(* IEC 61131-3 sources: plc-st-coding-agent/progress/evidence/f14_v2_public_20261112b/jobs/codex_deepseek-v4pro, 5 files *)

(* ---- public-easy-01.candidate_01.st ---- *)
FUNCTION_BLOCK FillingLineControl
VAR_INPUT
    bottleSensor : BOOL;
    cleaningConfirmButton : BOOL;
    fillingConfirmButton : BOOL;
    cappingConfirmButton : BOOL;
    packingConfirmButton : BOOL;
    finishedButton : BOOL;
END_VAR
VAR_OUTPUT
    Pump_Motor : BOOL;
    Filling_Valve : BOOL;
    Capping_Machine : BOOL;
    Packing_Machine : BOOL;
    Completion_Light : BOOL;
END_VAR
VAR
    step : INT := 0;
END_VAR

CASE step OF
    0:
        IF bottleSensor THEN
            step := 1;
        END_IF;

    1:
        IF cleaningConfirmButton THEN
            step := 2;
        END_IF;

    2:
        IF fillingConfirmButton THEN
            step := 3;
        END_IF;

    3:
        IF cappingConfirmButton THEN
            step := 4;
        END_IF;

    4:
        IF packingConfirmButton THEN
            step := 5;
        END_IF;

    5:
        IF finishedButton THEN
            step := 0;
        END_IF;
END_CASE;

Pump_Motor := (step = 1);
Filling_Valve := (step = 2);
Capping_Machine := (step = 3);
Packing_Machine := (step = 4);
Completion_Light := (step = 5);

END_FUNCTION_BLOCK

(* ---- public-easy-02.candidate_01.st ---- *)
FUNCTION_BLOCK FB
VAR_INPUT
    value : DWORD;
END_VAR
VAR_OUTPUT
    hasChanged : BOOL;
    hasRisingEdges : BOOL;
    risingBits : DWORD;
    noOfRisingBits : USINT;
    hasFallingEdges : BOOL;
    fallingBits : DWORD;
    noOfFallingBits : USINT;
END_VAR
VAR
    lastValue : DWORD;
    firstCycle : BOOL := TRUE;
    bitMask : DWORD;
    bitIndex : INT;
END_VAR

noOfRisingBits := USINT#0;
noOfFallingBits := USINT#0;

IF firstCycle THEN
    lastValue := value;
    firstCycle := FALSE;
    hasChanged := FALSE;
    hasRisingEdges := FALSE;
    risingBits := DWORD#0;
    hasFallingEdges := FALSE;
    fallingBits := DWORD#0;
ELSE
    hasChanged := (lastValue <> value);
    risingBits := (NOT lastValue) AND value;
    fallingBits := lastValue AND (NOT value);

    hasRisingEdges := (risingBits <> DWORD#0);
    hasFallingEdges := (fallingBits <> DWORD#0);

    FOR bitIndex := 0 TO 31 DO
        bitMask := SHL(DWORD#1, bitIndex);
        IF ((risingBits AND bitMask) <> DWORD#0) THEN
            noOfRisingBits := noOfRisingBits + USINT#1;
        END_IF;
        IF ((fallingBits AND bitMask) <> DWORD#0) THEN
            noOfFallingBits := noOfFallingBits + USINT#1;
        END_IF;
    END_FOR;

    lastValue := value;
END_IF;

END_FUNCTION_BLOCK

(* ---- public-easy-02.candidate_02.st ---- *)
FUNCTION_BLOCK FB
VAR_INPUT
    value : DWORD;
END_VAR
VAR_OUTPUT
    hasChanged : BOOL;
    hasRisingEdges : BOOL;
    risingBits : DWORD;
    noOfRisingBits : USINT;
    hasFallingEdges : BOOL;
    fallingBits : DWORD;
    noOfFallingBits : USINT;
END_VAR
VAR
    lastValue : DWORD;
    bitIndex : INT;
END_VAR

risingBits := (NOT lastValue) AND value;
fallingBits := lastValue AND (NOT value);

hasChanged := lastValue <> value;
hasRisingEdges := risingBits <> DWORD#0;
hasFallingEdges := fallingBits <> DWORD#0;

noOfRisingBits := USINT#0;
noOfFallingBits := USINT#0;

FOR bitIndex := 0 TO 31 DO
    IF ((SHR(risingBits, bitIndex) AND DWORD#1) <> DWORD#0) THEN
        noOfRisingBits := noOfRisingBits + USINT#1;
    END_IF;

    IF ((SHR(fallingBits, bitIndex) AND DWORD#1) <> DWORD#0) THEN
        noOfFallingBits := noOfFallingBits + USINT#1;
    END_IF;
END_FOR;

lastValue := value;

END_FUNCTION_BLOCK

(* ---- public-easy-03.candidate_01.st ---- *)
FUNCTION_BLOCK AlarmHandling
VAR_INPUT
    Value : REAL;
    hiLevel : REAL;
    loLevel : REAL;
    hystWindow : REAL;
END_VAR

VAR_OUTPUT
    hiAlarm : BOOL;
    loAlarm : BOOL;
    error : BOOL;
    status : WORD;
END_VAR

VAR
    hiAlarmState : BOOL;
    loAlarmState : BOOL;
END_VAR

BEGIN
    hiAlarm := FALSE;
    loAlarm := FALSE;
    error := FALSE;
    status := 16#0000;

    IF loLevel >= hiLevel THEN
        error := TRUE;
        status := 16#8001;
        RETURN;
    END_IF;

    IF hystWindow >= (hiLevel - loLevel) THEN
        error := TRUE;
        status := 16#8002;
        RETURN;
    END_IF;

    IF Value > hiLevel THEN
        hiAlarmState := TRUE;
    ELSIF Value < (hiLevel - hystWindow) THEN
        hiAlarmState := FALSE;
    END_IF;

    IF Value < loLevel THEN
        loAlarmState := TRUE;
    ELSIF Value > (loLevel + hystWindow) THEN
        loAlarmState := FALSE;
    END_IF;

    hiAlarm := hiAlarmState;
    loAlarm := loAlarmState;
END_FUNCTION_BLOCK

(* ---- public-easy-03.candidate_02.st ---- *)
FUNCTION_BLOCK AlarmHandling
VAR_INPUT
    Value : REAL;
    hiLevel : REAL;
    loLevel : REAL;
    hystWindow : REAL;
END_VAR

VAR_OUTPUT
    hiAlarm : BOOL;
    loAlarm : BOOL;
    error : BOOL;
    status : WORD;
END_VAR

BEGIN
    error := FALSE;
    status := WORD#16#0000;

    IF loLevel >= hiLevel THEN
        hiAlarm := FALSE;
        loAlarm := FALSE;
        error := TRUE;
        status := WORD#16#8001;
    ELSIF hystWindow >= (hiLevel - loLevel) THEN
        hiAlarm := FALSE;
        loAlarm := FALSE;
        error := TRUE;
        status := WORD#16#8002;
    ELSE
        IF Value > hiLevel THEN
            hiAlarm := TRUE;
        ELSIF Value < (hiLevel - hystWindow) THEN
            hiAlarm := FALSE;
        END_IF;

        IF Value < loLevel THEN
            loAlarm := TRUE;
        ELSIF Value > (loLevel + hystWindow) THEN
            loAlarm := FALSE;
        END_IF;
    END_IF;
END_FUNCTION_BLOCK
